// TIA Portal V21 export
// export: Created 2026-11-10T07:35:05.8371291Z, ExportSetting WithDefaults, DisplayName Totally Integrated Automation Portal, DisplayVersion V21 Update 3, DisplayName STEP 7 Professional, DisplayVersion V21 Update 3, DisplayName STEP 7 Safety, DisplayVersion V21, DisplayName Tech WebApplication, DisplayVersion V21, DisplayName WinCC Basic/Comfort/Advanced, DisplayVersion V21 Update 3, DisplayName WinCC Unified, DisplayVersion V21 Update 3
FUNCTION_BLOCK "FB_Lad_ex047"   // FB92, LAD
{ S7_Optimized_Access := 'TRUE' }
VERSION : 0.1
// stored: AutoNumber true, IsIECCheckEnabled false, IsRetainMemResEnabled false, MemoryReserve 100, SetENOAutomatically false, UDAEnableTagReadback false
   VAR_INPUT
      v_id : HW_SUBMODULE;
   END_VAR
   VAR_OUTPUT
      v_status : DWord;
      v_len : Int;
   END_VAR
   VAR_IN_OUT
      v_inputs : Array[0..99] of Byte;
   END_VAR
   VAR
      inst { S7_SetPoint := 'True'} : GETIO;
   END_VAR
BEGIN

REGION Network 1: GETIO - Read all inputs of a submodule
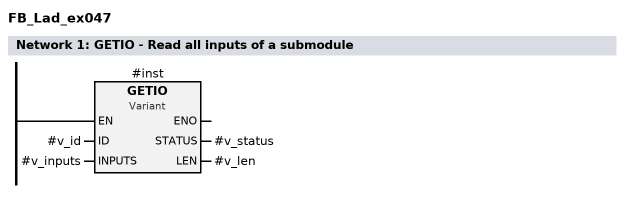
   RUNG wire#powerrail
      { S7_Templates := "[ptr_type := Variant, id_type := HW_SUBMODULE]" } #inst.GETIO(ID := #v_id, STATUS => #v_status, LEN => #v_len, INPUTS := #v_inputs)
   END_RUNG
   // the same network as SCL:
   #inst(ID := #v_id, INPUTS := #v_inputs, STATUS => #v_status, LEN => #v_len);   // GETIO
END_REGION
END_FUNCTION_BLOCK
